(* IEC 61131-3 sources: moqui-plc/codesys-v4/moqui-plc.fbsdev/moqui.iecapp^/moqui/framework/src/test/context, 1 file *)

(* ---- LogTestSuite.prg.st ---- *)
(*
 * Log pipeline test suite: LogRingBuffer, LoggerFacade registration, level threshold, duplicate summaries
 * and rate limit.
 * It runs once; passed is TRUE when every check holds, otherwise failedCheck is the number of the first failed check.
 *
 * Run it in its own test task with MqttCommunication not running: the suite reads the registered buffer itself,
 * and LogDispatcher would otherwise publish and release the test records.
 *)
PROGRAM LogTestSuite

	VAR
		finished : BOOL;
		passed : BOOL;
		checks : UINT;
		failedCheck : UINT;
		ring : LogRingBuffer;
		facade : LoggerFacade;
		limitedFacade : LoggerFacade;
		event : LogEvent;
		source : REFERENCE TO LogSource;
		savedMinLevel : LogLevel;
		writtenBefore : DINT;
		i : UINT;
		previous : DINT;
		ok : BOOL;
	END_VAR

	IF finished THEN RETURN; END_IF;
	finished := TRUE;
	passed := TRUE;

	(* ========== LogRingBuffer: fills, refuses without overwriting, accepts again once released ========== *)
	event.loggerName := 'LOG_TEST';
	event.payloadType := LogPayloadType.Text;
	event.payload.message := 'ring';
	ok := TRUE;
	FOR i := 1 TO MoquiConf.LOG_MAX_SIZE DO
		ring(cmd := LogCmd.Push, logEntry := event);
		ok := ok AND ring.done AND NOT ring.dropped;
	END_FOR;
	checks := checks + 1; IF NOT ok AND (failedCheck = 0) THEN failedCheck := checks; END_IF;
	checks := checks + 1; IF NOT ring.isFull AND (failedCheck = 0) THEN failedCheck := checks; END_IF;

	ring(cmd := LogCmd.Push, logEntry := event);
	checks := checks + 1; IF NOT (ring.dropped AND (ring.droppedCount = 1) AND NOT ring.done) AND (failedCheck = 0) THEN failedCheck := checks; END_IF;
	checks := checks + 1; IF NOT ((ring.logBuffer[1].sequence = 1) AND (ring.logBuffer[MoquiConf.LOG_MAX_SIZE].sequence = MoquiConf.LOG_MAX_SIZE))
			AND (failedCheck = 0) THEN failedCheck := checks; END_IF;

	(* The consumer releases one record: its slot is reused by the next record *)
	previous := __XADD(ADR(ring.readCount), 1);
	ring(cmd := LogCmd.Push, logEntry := event);
	checks := checks + 1; IF NOT (ring.done AND (ring.logBuffer[1].sequence = UINT_TO_UDINT(MoquiConf.LOG_MAX_SIZE) + 1))
			AND (failedCheck = 0) THEN failedCheck := checks; END_IF;
	checks := checks + 1; IF NOT ((ring.writeCount - ring.readCount) = UINT_TO_DINT(MoquiConf.LOG_MAX_SIZE)) AND (failedCheck = 0) THEN failedCheck := checks; END_IF;

	(* ========== LoggerFacade: registration, level threshold, duplicate summary ========== *)
	savedMinLevel := ec.logMinLevel;
	ec.logMinLevel := LogLevel.Info;

	facade.enable := TRUE;
	facade.loggerName := 'LOG_TEST';
	facade.level := LogLevel.Info;
	facade.suppressDuplicates := TRUE;
	facade.suppressDuration := T#1H;

	facade(message := 'first');
	checks := checks + 1; IF NOT (facade.done AND NOT facade.error) AND (failedCheck = 0) THEN failedCheck := checks; END_IF;
	checks := checks + 1; IF NOT ((ec.logSourceListSize >= 1) AND (ec.logSourceListSize <= UINT_TO_DINT(MoquiConf.LOG_SOURCE_LIST_MAX_SIZE)))
			AND (failedCheck = 0) THEN failedCheck := checks; END_IF;

	IF failedCheck = 0 THEN
		source REF= ec.logSourceList[DINT_TO_UINT(ec.logSourceListSize)];
		writtenBefore := source.logRef.writeCount;

		(* Two repetitions are only counted *)
		facade(message := 'first');
		facade(message := 'first');
		checks := checks + 1; IF NOT (facade.done AND (source.logRef.writeCount = writtenBefore)) AND (failedCheck = 0) THEN failedCheck := checks; END_IF;

		(* A Debug event is below the threshold *)
		facade(message := 'debug', level := LogLevel.Debug);
		checks := checks + 1; IF NOT (NOT facade.done AND (source.logRef.writeCount = writtenBefore)) AND (failedCheck = 0) THEN failedCheck := checks; END_IF;

		(* A different event writes the summary of the repetitions, then itself *)
		facade(message := 'second', level := LogLevel.Info);
		checks := checks + 1; IF NOT (source.logRef.writeCount = writtenBefore + 2) AND (failedCheck = 0) THEN failedCheck := checks; END_IF;
		checks := checks + 1; IF NOT ((source.logRef.logBuffer[2].repeatCount = 2) AND (source.logRef.logBuffer[2].payload.message = 'first')
				AND (source.logRef.logBuffer[3].repeatCount = 1) AND (source.logRef.logBuffer[3].payload.message = 'second'))
				AND (failedCheck = 0) THEN failedCheck := checks; END_IF;
		checks := checks + 1; IF NOT ((source.logRef.logBuffer[1].sequence = 1) AND (source.logRef.logBuffer[3].sequence = 3))
				AND (failedCheck = 0) THEN failedCheck := checks; END_IF;
	END_IF;

	(* ========== LoggerFacade: rate limit with alternating events ========== *)
	limitedFacade.enable := TRUE;
	limitedFacade.loggerName := 'LOG_RATE_TEST';
	limitedFacade.level := LogLevel.Info;
	limitedFacade.suppressDuplicates := TRUE;
	limitedFacade.suppressDuration := T#1H;
	limitedFacade.maxEventsPerWindow := 3;

	limitedFacade(message := 'a');
	IF failedCheck = 0 THEN
		source REF= ec.logSourceList[DINT_TO_UINT(ec.logSourceListSize)];
		writtenBefore := source.logRef.writeCount;

		(* 'b' and 'a' fill the window (3 events), then the alternation is only counted: no summary per call *)
		FOR i := 1 TO 10 DO
			limitedFacade(message := 'b');
			limitedFacade(message := 'a');
		END_FOR;
		checks := checks + 1; IF NOT (source.logRef.writeCount = writtenBefore + 2) AND (failedCheck = 0) THEN failedCheck := checks; END_IF;

		limitedFacade(message := 'b');
		checks := checks + 1; IF NOT (limitedFacade.rateLimited AND NOT limitedFacade.done
				AND (source.logRef.writeCount = writtenBefore + 2)) AND (failedCheck = 0) THEN failedCheck := checks; END_IF;
	END_IF;

	ec.logMinLevel := savedMinLevel;
	passed := failedCheck = 0;
	END_PROGRAM
